KUKA KRL program: bt_sps.src

&ACCESS RVP
&REL 1
&COMMENT bt2krl sim submit part plan 16#F77E
DEF BT_SPS()
   DECL INT BT_Q
   DECL BOOL BT_PRUN
   ; Generated by bt2krl 0.1.0 from bt2plc plan bt_1790934549_welding_cell_2_small (cell welding_cell_2_small), PLAN_ID 16#F77E
   ; Robot robot1 (R1), controller robot1, model KR240R2900_ULTRA, joint mapping identity
   ; Profile sim (bt2plc simulator telegram). NEVER install on a VW KS24 robot:
   ; its signals collide with the VW standard (Fertigmeldung, interlocks, PRG_NR).
   ; Do not edit: regenerate with bt2krl (plain KRL, no inline forms).
   ; Call once per cycle from the LOOP of KRC/R1/System/sps.sub (fold USER PLC): BT_SPS()
   ; Job handshake as the bt2plc device simulator (FB_VASS_DeviceSimulator).
   ;FOLD READY AND ABORT
      BT_READY=$PERI_RDY AND ($MODE_OP==#EX) AND NOT BT_ERR AND NOT (BT_RUN AND NOT BT_ABRT) AND $ALARM_STOP AND $USER_SAF
      IF BT_RUN AND NOT BT_ABRT THEN
         IF BT_C_STOP OR BT_C_CANCEL OR NOT $PERI_RDY OR NOT $ALARM_STOP OR ($PRO_STATE1<>#P_ACTIVE) THEN
            BT_ABRT=TRUE
         ENDIF
      ENDIF
   ;ENDFOLD
   ;FOLD JOB HANDSHAKE
      IF BT_C_JOBREQ AND NOT BT_M_JOB AND BT_READY THEN
         BT_JOBNR=BT_JOB
         BT_PLANL=BT_PLANID
         BT_ACK=TRUE
         BT_FIN=FALSE
      ENDIF
      IF NOT BT_C_JOBREQ THEN
         BT_ACK=FALSE
      ENDIF
      BT_M_JOB=BT_C_JOBREQ
      IF BT_C_START AND NOT BT_M_START AND BT_READY AND (BT_JOBNR<>0) THEN
         BT_START=TRUE
      ENDIF
      BT_M_START=BT_C_START
   ;ENDFOLD
   ;FOLD RESET: edge clears the warning, held 500 ms clears the error
      IF BT_C_RESET THEN
         IF NOT BT_M_RESET THEN
            BT_WCODE=0
            $TIMER[20]=0
            $TIMER_STOP[20]=FALSE
         ENDIF
         IF BT_ERR AND ($TIMER[20]>=500) THEN
            BT_ERR=FALSE
            BT_ECODE=0
            BT_WCODE=0
         ENDIF
      ELSE
         $TIMER_STOP[20]=TRUE
      ENDIF
      BT_M_RESET=BT_C_RESET
   ;ENDFOLD
   ;FOLD NO FOLGE ACTIVE: STEP := 0, REQUEST := 0 (outputs persist after a cancel)
      IF NOT BT_RUN OR BT_ABRT THEN
         BT_STEP=0
         BT_REQ0=0
         BT_REQ1=0
         BT_REQ2=0
         BT_REQ3=0
      ENDIF
   ;ENDFOLD
   ;FOLD STATUS
      ; ProgRunning low only after ProgFinished is out: read BT_RUN first, write BT_O_FIN first
      BT_PRUN=BT_RUN AND NOT BT_ABRT
      BT_O_FIN=BT_FIN
      BT_O_RUN=BT_PRUN
      BT_O_DRIVES=$PERI_RDY
      BT_O_HOME=(ABS($AXIS_ACT.A1-BT_HOME.A1)<=0.5) AND (ABS($AXIS_ACT.A2-BT_HOME.A2)<=0.5) AND (ABS($AXIS_ACT.A3-BT_HOME.A3)<=0.5) AND (ABS($AXIS_ACT.A4-BT_HOME.A4)<=0.5) AND (ABS($AXIS_ACT.A5-BT_HOME.A5)<=0.5) AND (ABS($AXIS_ACT.A6-BT_HOME.A6)<=0.5)
      BT_O_INPOS=NOT BT_RUN
      BT_O_EXT=($MODE_OP==#EX)
      BT_O_READY=BT_READY
      BT_O_ERROR=BT_ERR
      BT_O_WARN=(BT_WCODE<>0)
      BT_O_GATES=$USER_SAF
      BT_O_ESTOP=$ALARM_STOP
      BT_O_JOBACK=BT_ACK
      BT_O_PERIPH=TRUE
      BT_ECHO=BT_JOBNR
      BT_ERRCODE=BT_ECODE
      BT_WARNCODE=BT_WCODE
   ;ENDFOLD
   ;FOLD JOINT ENCODER: A1..A6 as INT16 big-endian, 0.02 deg/count, bytes 16-27
      BT_Q=$AXIS_ACT.A1*50
      IF BT_Q<0 THEN
         BT_Q=BT_Q+65536
      ENDIF
      BT_JNT0=(BT_Q-(BT_Q B_AND 255))/256
      BT_JNT1=BT_Q B_AND 255
      BT_Q=$AXIS_ACT.A2*50
      IF BT_Q<0 THEN
         BT_Q=BT_Q+65536
      ENDIF
      BT_JNT2=(BT_Q-(BT_Q B_AND 255))/256
      BT_JNT3=BT_Q B_AND 255
      BT_Q=$AXIS_ACT.A3*50
      IF BT_Q<0 THEN
         BT_Q=BT_Q+65536
      ENDIF
      BT_JNT4=(BT_Q-(BT_Q B_AND 255))/256
      BT_JNT5=BT_Q B_AND 255
      BT_Q=$AXIS_ACT.A4*50
      IF BT_Q<0 THEN
         BT_Q=BT_Q+65536
      ENDIF
      BT_JNT6=(BT_Q-(BT_Q B_AND 255))/256
      BT_JNT7=BT_Q B_AND 255
      BT_Q=$AXIS_ACT.A5*50
      IF BT_Q<0 THEN
         BT_Q=BT_Q+65536
      ENDIF
      BT_JNT8=(BT_Q-(BT_Q B_AND 255))/256
      BT_JNT9=BT_Q B_AND 255
      BT_Q=$AXIS_ACT.A6*50
      IF BT_Q<0 THEN
         BT_Q=BT_Q+65536
      ENDIF
      BT_JNT10=(BT_Q-(BT_Q B_AND 255))/256
      BT_JNT11=BT_Q B_AND 255
   ;ENDFOLD
END
